(* IEC 61131-3 sources: freecad-ai-parts/factory/digital/vplc/examples, 2 files *)

(* ---- press_p15_5_1.st ---- *)
(* 程序 15.5.1  压装工位：加上异常处理——动作超时、传感器冲突、急停与恢复 *)
TYPE E_Press : (INIT, HOMING, IDLE, CLAMPING, PRESSING, RETURNING, UNCLAMPING, FAULT, ESTOP); END_TYPE

PROGRAM Main
  VAR
    state : E_Press := INIT;
    prev : E_Press := INIT;    (* 上一次扫描的状态：状态一变，计时重新开始 *)
    tState : TON;              (* 本状态已经停留的时间 *)
    maxTime : TIME;            (* 本状态允许停留的最长时间 *)
    faultCode : INT;               (* 故障代码：0 无；1 夹紧超时；2 压装超时；3 回程超时；4 松开超时；5 回原点超时；9 传感器冲突 *)
    clampHold : BOOL;          (* 进入故障或急停时夹具是否夹着：保持原样 *)
    auto, go, jog : BOOL;
    rStep, rReset : R_TRIG;
    tTwoHand : TON;
    force, peak : REAL;
    resOk, resNok : BOOL;
  END_VAR

  force := INT_TO_REAL(AI_Force) * 10.0 / 27648.0;
  tTwoHand(IN := S_Hand1 OR S_Hand2, PT := T#500ms);
  rStep(CLK := S_Step);
  rReset(CLK := S_Reset);
  auto := S_Auto;
  go := auto OR rStep.Q;

  (* 1. 急停与传感器冲突：任何状态下都优先 *)
  IF NOT S_EStop AND state <> ESTOP THEN
    clampHold := Y_Clamp; state := ESTOP;
  ELSIF ((B_Clamped AND B_Unclamped) OR (B_PressUp AND B_PressDown)) AND state <> FAULT AND state <> ESTOP THEN
    clampHold := Y_Clamp; faultCode := 9; state := FAULT;
  END_IF;

  (* 2. 状态时限：自动方式和回原点时才计时（单步时等的是人） *)
  CASE state OF
    CLAMPING, UNCLAMPING: maxTime := T#1s;
    PRESSING: maxTime := T#4s;
    RETURNING: maxTime := T#5s;
    HOMING: maxTime := T#5s;
  ELSE
    maxTime := T#1h;
  END_CASE;
  tState(IN := state = prev AND (auto OR state = HOMING), PT := maxTime);
  prev := state;

  (* 3. 转移 *)
  CASE state OF
    INIT:
      IF rReset.Q THEN state := HOMING; END_IF;
    HOMING:
      IF B_PressUp AND B_Unclamped THEN state := IDLE;
      ELSIF tState.Q THEN clampHold := FALSE; faultCode := 5; state := FAULT; END_IF;
    IDLE:
      IF rReset.Q THEN
        state := HOMING;
      ELSIF B_Part AND B_PressUp AND B_Unclamped AND S_LC
            AND ((auto AND S_Hand1 AND S_Hand2 AND NOT tTwoHand.Q) OR (NOT auto AND rStep.Q)) THEN
        resOk := FALSE; resNok := FALSE; peak := 0.0;
        state := CLAMPING;
      ELSIF NOT auto AND (S_JogClamp OR S_JogDown OR S_JogUp) THEN
        state := INIT;                    (* 点动过：位置不再确定，再启动前要回原点 *)
      END_IF;
    CLAMPING:
      IF go AND B_Clamped THEN state := PRESSING;
      ELSIF tState.Q THEN clampHold := TRUE; faultCode := 1; state := FAULT; END_IF;
    PRESSING:
      peak := MAX(peak, force);
      IF force > 8.0 THEN
        resNok := TRUE; state := RETURNING;
      ELSIF go AND B_PressDown THEN
        resOk := peak >= 4.0 AND peak <= 7.0; resNok := NOT resOk;
        state := RETURNING;
      ELSIF auto AND NOT (S_Hand1 AND S_Hand2 AND S_LC) THEN
        resNok := TRUE; state := RETURNING;
      ELSIF tState.Q THEN clampHold := TRUE; faultCode := 2; state := FAULT; END_IF;
    RETURNING:
      IF go AND B_PressUp THEN state := UNCLAMPING;
      ELSIF tState.Q THEN clampHold := TRUE; faultCode := 3; state := FAULT; END_IF;
    UNCLAMPING:
      IF go AND B_Unclamped THEN state := IDLE;
      ELSIF tState.Q THEN clampHold := FALSE; faultCode := 4; state := FAULT; END_IF;
    FAULT:                                (* 停在原地，等人看清原因、按复位 *)
      IF rReset.Q AND S_EStop AND NOT ((B_Clamped AND B_Unclamped) OR (B_PressUp AND B_PressDown)) THEN
        faultCode := 0; state := HOMING;
      END_IF;
    ESTOP:                                (* 急停松开后也不自己动，按复位才回原点 *)
      IF S_EStop AND rReset.Q THEN state := HOMING; END_IF;
  END_CASE;

  (* 4. 输出 *)
  jog := NOT auto AND (state = IDLE OR state = INIT OR state = FAULT);   (* 故障时允许点动，联锁照样有效 *)
  Y_Clamp     := state = CLAMPING OR state = PRESSING OR state = RETURNING OR (jog AND S_JogClamp)
                 OR ((state = FAULT OR state = ESTOP) AND clampHold);
  Y_PressDown := ((state = PRESSING AND S_Hand1 AND S_Hand2) OR (jog AND S_JogDown AND B_Clamped)) AND S_LC AND S_EStop;
  Y_PressUp   := (state = RETURNING OR (state = HOMING AND NOT B_PressUp) OR (jog AND S_JogUp))
                 AND S_EStop AND NOT Y_PressDown;
  H_OK    := resOk;
  H_NOK   := resNok;
  H_Ready := state = IDLE;
  H_Fault := state = FAULT OR state = ESTOP;
END_PROGRAM

(* ---- sorter_ref.st ---- *)
(* 数字工厂分拣线 SORT-01 的参考程序：先进先出跟踪分拣（金属 → 1 号箱，红 → 2 号箱，蓝 → 3 号箱，高件 → 末端废品），
   推杆伸出 0.3 s 不到位即报故障（faultCode = 推杆号）：输送带停、故障灯亮；按停止再按启动恢复，带上剩下的件放行到末端。 *)
PROGRAM Main
  VAR
    kind : ARRAY[0..31] OF INT;          (* 1 金属 2 红 3 蓝 9 废品（高件） *)
    gone : ARRAY[0..31] OF BOOL;
    nIn, s1, s2, s3 : INT;               (* 进检测工位的件数；各推杆已处理到第几件 *)
    rIn, r1, r2, r3, rStart : R_TRIG;
    push1, push2, push3 : TP;
    t1, t2, t3 : TON;                    (* 推杆伸出监视 *)
    run, fault : BOOL;
    faultCode : INT;
    k : INT;
  END_VAR

  (* 启停与故障复位：停止（常闭）断开即复位故障；启动的上升沿重新开始，带上的件不再跟踪 *)
  rStart(CLK := S_Start);
  IF NOT S_Stop THEN fault := FALSE; faultCode := 0; END_IF;
  IF rStart.Q AND S_Stop AND NOT fault THEN run := TRUE; s1 := nIn; s2 := nIn; s3 := nIn; END_IF;
  IF NOT S_Stop OR fault THEN run := FALSE; END_IF;

  (* 检测工位：记下这一件该去哪里 *)
  rIn(CLK := B_Insp);
  IF rIn.Q AND run THEN
    IF B_Tall THEN k := 9; ELSIF B_Metal THEN k := 1; ELSIF B_Red THEN k := 2; ELSE k := 3; END_IF;
    kind[nIn MOD 32] := k; gone[nIn MOD 32] := FALSE; nIn := nIn + 1;
  END_IF;

  (* 三个推杆：件到了推杆前，按队列里的记录决定推不推 *)
  r1(CLK := B_P1);
  IF r1.Q AND s1 < nIn THEN
    IF kind[s1 MOD 32] = 1 THEN gone[s1 MOD 32] := TRUE; push1(IN := TRUE, PT := T#400ms); END_IF;
    s1 := s1 + 1;
  END_IF;
  r2(CLK := B_P2);
  IF r2.Q THEN
    WHILE s2 < nIn AND gone[s2 MOD 32] AND s2 < s1 DO s2 := s2 + 1; END_WHILE;
    IF s2 < nIn THEN IF kind[s2 MOD 32] = 2 THEN gone[s2 MOD 32] := TRUE; push2(IN := TRUE, PT := T#400ms); END_IF; s2 := s2 + 1; END_IF;
  END_IF;
  r3(CLK := B_P3);
  IF r3.Q THEN
    WHILE s3 < nIn AND gone[s3 MOD 32] AND s3 < s2 DO s3 := s3 + 1; END_WHILE;
    IF s3 < nIn THEN IF kind[s3 MOD 32] = 3 THEN gone[s3 MOD 32] := TRUE; push3(IN := TRUE, PT := T#400ms); END_IF; s3 := s3 + 1; END_IF;
  END_IF;
  push1(IN := FALSE); push2(IN := FALSE); push3(IN := FALSE);

  (* 推杆监视：电磁阀得电 0.3 s 还没伸出到位，就是推杆卡住或到位开关坏了 *)
  t1(IN := push1.Q AND NOT B_Y1Out, PT := T#300ms);
  t2(IN := push2.Q AND NOT B_Y2Out, PT := T#300ms);
  t3(IN := push3.Q AND NOT B_Y3Out, PT := T#300ms);
  IF NOT fault THEN
    IF t1.Q THEN fault := TRUE; faultCode := 1;
    ELSIF t2.Q THEN fault := TRUE; faultCode := 2;
    ELSIF t3.Q THEN fault := TRUE; faultCode := 3; END_IF;
  END_IF;

  M_Belt := run AND NOT fault;
  Y1 := push1.Q AND NOT fault;
  Y2 := push2.Q AND NOT fault;
  Y3 := push3.Q AND NOT fault;
  H_Run := run;
  H_Fault := fault;
END_PROGRAM
